(* IEC 61131-3 sources: rusty/tests/lit/single/type_promotion/case_selector, 7 files *)

(* ---- derived_selector_range_across_midpoint.st ---- *)
// RUN: %COMPILE %s && %RUN | %CHECK %s
// A range label that crosses the signed midpoint matches every value between its bounds, also through an alias or subrange type.
TYPE
    Level : USINT;
    Small : UINT(0..60000);
END_TYPE

FUNCTION branch_alias : DINT
    VAR_INPUT
        x : Level;
    END_VAR

    CASE x OF
        100..200: branch_alias := 1;
    ELSE
        branch_alias := 9;
    END_CASE
END_FUNCTION

FUNCTION branch_subrange : DINT
    VAR_INPUT
        x : Small;
    END_VAR

    CASE x OF
        30000..50000: branch_subrange := 1;
    ELSE
        branch_subrange := 9;
    END_CASE
END_FUNCTION

FUNCTION branch_list : DINT
    VAR_INPUT
        x : USINT;
    END_VAR

    CASE x OF
        1, 100..200, 250: branch_list := 1;
    ELSE
        branch_list := 9;
    END_CASE
END_FUNCTION

FUNCTION main : DINT
    printf('alias 150 -> %d$N', branch_alias(150));             // CHECK: alias 150 -> 1
    printf('subrange 40000 -> %d$N', branch_subrange(40000));   // CHECK-NEXT: subrange 40000 -> 1
    printf('list 1 -> %d$N', branch_list(1));                   // CHECK-NEXT: list 1 -> 1
    printf('list 150 -> %d$N', branch_list(150));               // CHECK-NEXT: list 150 -> 1
    printf('list 250 -> %d$N', branch_list(250));               // CHECK-NEXT: list 250 -> 1
END_FUNCTION

(* ---- signed_range_across_zero.st ---- *)
// RUN: %COMPILE %s && %RUN | %CHECK %s
// Range labels that cross zero on a signed selector.
FUNCTION branch_sint : DINT
    VAR_INPUT
        x : SINT;
    END_VAR

    CASE x OF
        -128..-100: branch_sint := 1;
        -10..10: branch_sint := 2;
        100..127: branch_sint := 3;
    ELSE
        branch_sint := 9;
    END_CASE
END_FUNCTION

FUNCTION branch_int : DINT
    VAR_INPUT
        x : INT;
    END_VAR

    CASE x OF
        -32768..-30000: branch_int := 1;
        -1000..1000: branch_int := 2;
    ELSE
        branch_int := 9;
    END_CASE
END_FUNCTION

FUNCTION branch_dint : DINT
    VAR_INPUT
        x : DINT;
    END_VAR

    CASE x OF
        -2147483648..-2000000000: branch_dint := 1;
        -1000000000..1000000000: branch_dint := 2;
    ELSE
        branch_dint := 9;
    END_CASE
END_FUNCTION

FUNCTION branch_lint : DINT
    VAR_INPUT
        x : LINT;
    END_VAR

    CASE x OF
        -9223372036854775807..-9000000000000000000: branch_lint := 1;
        -5000000000..5000000000: branch_lint := 2;
    ELSE
        branch_lint := 9;
    END_CASE
END_FUNCTION

FUNCTION main : DINT
    // SINT
    printf('SINT -128 -> %d$N', branch_sint(-128));         // CHECK: SINT -128 -> 1
    printf('SINT -5 -> %d$N', branch_sint(-5));             // CHECK-NEXT: SINT -5 -> 2
    printf('SINT 5 -> %d$N', branch_sint(5));               // CHECK-NEXT: SINT 5 -> 2
    printf('SINT 127 -> %d$N', branch_sint(127));           // CHECK-NEXT: SINT 127 -> 3
    printf('SINT -50 -> %d$N', branch_sint(-50));           // CHECK-NEXT: SINT -50 -> 9

    // INT
    printf('INT -32768 -> %d$N', branch_int(-32768));       // CHECK-NEXT: INT -32768 -> 1
    printf('INT -500 -> %d$N', branch_int(-500));           // CHECK-NEXT: INT -500 -> 2
    printf('INT 2000 -> %d$N', branch_int(2000));           // CHECK-NEXT: INT 2000 -> 9

    // DINT
    printf('DINT -2147483648 -> %d$N', branch_dint(-2147483648));   // CHECK-NEXT: DINT -2147483648 -> 1
    printf('DINT -7 -> %d$N', branch_dint(-7));                     // CHECK-NEXT: DINT -7 -> 2

    // LINT
    printf('LINT -9100000000000000000 -> %d$N', branch_lint(-9100000000000000000));    // CHECK-NEXT: LINT -9100000000000000000 -> 1
    printf('LINT -4000000000 -> %d$N', branch_lint(-4000000000));                      // CHECK-NEXT: LINT -4000000000 -> 2
END_FUNCTION

(* ---- udint_range_across_midpoint.st ---- *)
// RUN: %COMPILE %s && %RUN | %CHECK %s
// A range label that crosses the signed midpoint of the UDINT selector matches every value between its bounds.
FUNCTION branch : DINT
    VAR_INPUT
        x : UDINT;
    END_VAR

    CASE x OF
        0:
            branch := 1;
        1..9:
            branch := 2;
        11..4294967294:
            branch := 3;
        4294967295:
            branch := 4;
    ELSE
        branch := 9;
    END_CASE
END_FUNCTION

FUNCTION main : DINT
    printf('0 -> %d$N', branch(0));                             // CHECK: 0 -> 1
    printf('5 -> %d$N', branch(5));                             // CHECK-NEXT: 5 -> 2
    printf('10 -> %d$N', branch(10));                           // CHECK-NEXT: 10 -> 9
    printf('11 -> %d$N', branch(11));                           // CHECK-NEXT: 11 -> 3
    printf('2147483647 -> %d$N', branch(2147483647));           // CHECK-NEXT: 2147483647 -> 3
    printf('2147483648 -> %d$N', branch(2147483648));           // CHECK-NEXT: 2147483648 -> 3
    printf('3000000000 -> %d$N', branch(3000000000));           // CHECK-NEXT: 3000000000 -> 3
    printf('4294967294 -> %d$N', branch(4294967294));           // CHECK-NEXT: 4294967294 -> 3
    printf('4294967295 -> %d$N', branch(4294967295));           // CHECK-NEXT: 4294967295 -> 4
END_FUNCTION

(* ---- uint_range_across_midpoint.st ---- *)
// RUN: %COMPILE %s && %RUN | %CHECK %s
// A range label that crosses the signed midpoint of the UINT selector matches every value between its bounds.
FUNCTION branch : DINT
    VAR_INPUT
        x : UINT;
    END_VAR

    CASE x OF
        0:
            branch := 1;
        1..9:
            branch := 2;
        11..65534:
            branch := 3;
        65535:
            branch := 4;
    ELSE
        branch := 9;
    END_CASE
END_FUNCTION

FUNCTION main : DINT
    printf('0 -> %d$N', branch(0));                             // CHECK: 0 -> 1
    printf('5 -> %d$N', branch(5));                             // CHECK-NEXT: 5 -> 2
    printf('10 -> %d$N', branch(10));                           // CHECK-NEXT: 10 -> 9
    printf('11 -> %d$N', branch(11));                           // CHECK-NEXT: 11 -> 3
    printf('32767 -> %d$N', branch(32767));                     // CHECK-NEXT: 32767 -> 3
    printf('32768 -> %d$N', branch(32768));                     // CHECK-NEXT: 32768 -> 3
    printf('40000 -> %d$N', branch(40000));                     // CHECK-NEXT: 40000 -> 3
    printf('65534 -> %d$N', branch(65534));                     // CHECK-NEXT: 65534 -> 3
    printf('65535 -> %d$N', branch(65535));                     // CHECK-NEXT: 65535 -> 4
END_FUNCTION

(* ---- ulint_range_across_midpoint.st ---- *)
// RUN: %COMPILE %s && %RUN | %CHECK %s
// A range label that crosses the signed midpoint of the ULINT selector matches every value between its bounds.
FUNCTION branch : DINT
    VAR_INPUT
        x : ULINT;
    END_VAR

    CASE x OF
        0:
            branch := 1;
        1..9:
            branch := 2;
        11..18446744073709551614:
            branch := 3;
        18446744073709551615:
            branch := 4;
    ELSE
        branch := 9;
    END_CASE
END_FUNCTION

FUNCTION main : DINT
    printf('0 -> %d$N', branch(0));                             // CHECK: 0 -> 1
    printf('5 -> %d$N', branch(5));                             // CHECK-NEXT: 5 -> 2
    printf('10 -> %d$N', branch(10));                           // CHECK-NEXT: 10 -> 9
    printf('11 -> %d$N', branch(11));                           // CHECK-NEXT: 11 -> 3
    printf('9223372036854775807 -> %d$N', branch(9223372036854775807));  // CHECK-NEXT: 9223372036854775807 -> 3
    printf('9223372036854775808 -> %d$N', branch(9223372036854775808));  // CHECK-NEXT: 9223372036854775808 -> 3
    printf('12000000000000000000 -> %d$N', branch(12000000000000000000));  // CHECK-NEXT: 12000000000000000000 -> 3
    printf('18446744073709551614 -> %d$N', branch(18446744073709551614));  // CHECK-NEXT: 18446744073709551614 -> 3
    printf('18446744073709551615 -> %d$N', branch(18446744073709551615));  // CHECK-NEXT: 18446744073709551615 -> 4
END_FUNCTION

(* ---- unsigned_range_within_one_half.st ---- *)
// RUN: %COMPILE %s && %RUN | %CHECK %s
// Range labels that stay below or above the signed midpoint of an unsigned selector.
FUNCTION branch_usint : DINT
    VAR_INPUT
        x : USINT;
    END_VAR

    CASE x OF
        1..100: branch_usint := 1;
        129..254: branch_usint := 2;
        255: branch_usint := 3;
    ELSE
        branch_usint := 9;
    END_CASE
END_FUNCTION

FUNCTION branch_uint : DINT
    VAR_INPUT
        x : UINT;
    END_VAR

    CASE x OF
        1..30000: branch_uint := 1;
        32769..65534: branch_uint := 2;
        65535: branch_uint := 3;
    ELSE
        branch_uint := 9;
    END_CASE
END_FUNCTION

FUNCTION branch_udint : DINT
    VAR_INPUT
        x : UDINT;
    END_VAR

    CASE x OF
        1..2000000000: branch_udint := 1;
        2147483649..4294967294: branch_udint := 2;
        4294967295: branch_udint := 3;
    ELSE
        branch_udint := 9;
    END_CASE
END_FUNCTION

FUNCTION branch_ulint : DINT
    VAR_INPUT
        x : ULINT;
    END_VAR

    CASE x OF
        1..9000000000000000000: branch_ulint := 1;
        9223372036854775809..18446744073709551614: branch_ulint := 2;
        18446744073709551615: branch_ulint := 3;
    ELSE
        branch_ulint := 9;
    END_CASE
END_FUNCTION

FUNCTION main : DINT
    // USINT
    printf('USINT 50 -> %d$N', branch_usint(50));                   // CHECK: USINT 50 -> 1
    printf('USINT 200 -> %d$N', branch_usint(200));                 // CHECK-NEXT: USINT 200 -> 2
    printf('USINT 255 -> %d$N', branch_usint(255));                 // CHECK-NEXT: USINT 255 -> 3
    printf('USINT 0 -> %d$N', branch_usint(0));                     // CHECK-NEXT: USINT 0 -> 9

    // UINT
    printf('UINT 100 -> %d$N', branch_uint(100));                   // CHECK-NEXT: UINT 100 -> 1
    printf('UINT 40000 -> %d$N', branch_uint(40000));               // CHECK-NEXT: UINT 40000 -> 2
    printf('UINT 65535 -> %d$N', branch_uint(65535));               // CHECK-NEXT: UINT 65535 -> 3

    // UDINT
    printf('UDINT 100 -> %d$N', branch_udint(100));                 // CHECK-NEXT: UDINT 100 -> 1
    printf('UDINT 3000000000 -> %d$N', branch_udint(3000000000));   // CHECK-NEXT: UDINT 3000000000 -> 2
    printf('UDINT 4294967295 -> %d$N', branch_udint(4294967295));   // CHECK-NEXT: UDINT 4294967295 -> 3

    // ULINT
    printf('ULINT 100 -> %d$N', branch_ulint(100));                 // CHECK-NEXT: ULINT 100 -> 1
    printf('ULINT 2^63 + 1 -> %d$N', branch_ulint(9223372036854775809));   // CHECK-NEXT: ULINT 2^63 + 1 -> 2
    printf('ULINT max -> %d$N', branch_ulint(18446744073709551615));       // CHECK-NEXT: ULINT max -> 3
END_FUNCTION

(* ---- usint_range_across_midpoint.st ---- *)
// RUN: %COMPILE %s && %RUN | %CHECK %s
// A range label that crosses the signed midpoint of the USINT selector matches every value between its bounds.
FUNCTION branch : DINT
    VAR_INPUT
        x : USINT;
    END_VAR

    CASE x OF
        0:
            branch := 1;
        1..9:
            branch := 2;
        11..254:
            branch := 3;
        255:
            branch := 4;
    ELSE
        branch := 9;
    END_CASE
END_FUNCTION

FUNCTION main : DINT
    printf('0 -> %d$N', branch(0));                             // CHECK: 0 -> 1
    printf('5 -> %d$N', branch(5));                             // CHECK-NEXT: 5 -> 2
    printf('10 -> %d$N', branch(10));                           // CHECK-NEXT: 10 -> 9
    printf('11 -> %d$N', branch(11));                           // CHECK-NEXT: 11 -> 3
    printf('127 -> %d$N', branch(127));                         // CHECK-NEXT: 127 -> 3
    printf('128 -> %d$N', branch(128));                         // CHECK-NEXT: 128 -> 3
    printf('200 -> %d$N', branch(200));                         // CHECK-NEXT: 200 -> 3
    printf('254 -> %d$N', branch(254));                         // CHECK-NEXT: 254 -> 3
    printf('255 -> %d$N', branch(255));                         // CHECK-NEXT: 255 -> 4
END_FUNCTION
